(* IEC 61131-3 sources: kns-port-domestic/targets/astra/lib/src/POUs/Util/FB_StartsWindow, 7 files *)

(* ---- FB_StartsWindow.decl.st ---- *)
// Назначение: пуски за скользящий час (лимит пусков двигателя). Кольцо отметок LTIME,
//             упорядоченных по времени: самая старая — в начале, самая новая — в конце.
//             Отметки старше окна и «из будущего» (время назад) удаляются. Окно не
//             энергонезависимо: после перезапуска ПЛК оно пустое (A-03).
// Автор:      kr0nsch
// Версия:     0.1.0
// Документ:   docs/fb/FB_StartsWindow.md
FUNCTION_BLOCK FB_StartsWindow
VAR
    altStart : ARRAY[0..GVL_Const.STARTS_WINDOW_MAX - 1] OF LTIME;   // кольцо отметок пусков
    uiNext   : UINT;      // индекс следующей записи
    uiUsed   : UINT;      // занято записей, 0..STARTS_WINDOW_MAX
END_VAR

(* ---- Count.method.decl.st ---- *)
// Число отметок t с t <= ltNow и ltNow - t < STARTS_WINDOW. Отметки «из будущего» (время
// назад) и старше окна удаляются
METHOD PUBLIC Count : UINT
VAR_INPUT
    ltNow : LTIME;    // текущее время
END_VAR
VAR
    xMore : BOOL;     // продолжать удаление
    uiLast : UINT;    // индекс самой новой отметки
    uiFirst : UINT;   // индекс самой старой отметки
END_VAR

(* ---- Count.method.impl.st ---- *)
// 1. Отметки «из будущего» — с конца
xMore := uiUsed > 0;
WHILE xMore DO
    uiLast := (uiNext + GVL_Const.STARTS_WINDOW_MAX - 1) MOD GVL_Const.STARTS_WINDOW_MAX;
    IF altStart[uiLast] > ltNow THEN
        uiNext := uiLast;
        uiUsed := uiUsed - 1;
        xMore := uiUsed > 0;
    ELSE
        xMore := FALSE;
    END_IF
END_WHILE

// 2. Отметки старше окна — с начала. Все оставшиеся <= ltNow: разность без переполнения
xMore := uiUsed > 0;
WHILE xMore DO
    uiFirst := (uiNext + GVL_Const.STARTS_WINDOW_MAX - uiUsed) MOD GVL_Const.STARTS_WINDOW_MAX;
    IF ltNow - altStart[uiFirst] >= GVL_Const.STARTS_WINDOW THEN
        uiUsed := uiUsed - 1;
        xMore := uiUsed > 0;
    ELSE
        xMore := FALSE;
    END_IF
END_WHILE

Count := uiUsed;

(* ---- Register.method.decl.st ---- *)
// Добавить отметку пуска; при заполнении кольца затирается самая старая
METHOD PUBLIC Register
VAR_INPUT
    ltNow : LTIME;   // время пуска
END_VAR
VAR
    xMore : BOOL;    // продолжать удаление с конца
    uiLast : UINT;   // индекс самой новой отметки
END_VAR

(* ---- Register.method.impl.st ---- *)
// 1. Отметки новее регистрируемой (было «время назад») удаляются: кольцо остаётся упорядоченным
xMore := uiUsed > 0;
WHILE xMore DO
    uiLast := (uiNext + GVL_Const.STARTS_WINDOW_MAX - 1) MOD GVL_Const.STARTS_WINDOW_MAX;
    IF altStart[uiLast] > ltNow THEN
        uiNext := uiLast;
        uiUsed := uiUsed - 1;
        xMore := uiUsed > 0;
    ELSE
        xMore := FALSE;
    END_IF
END_WHILE

// 2. Запись; заполненное кольцо затирает самую старую отметку
altStart[uiNext] := ltNow;
uiNext := (uiNext + 1) MOD GVL_Const.STARTS_WINDOW_MAX;
uiUsed := MIN(uiUsed + 1, GVL_Const.STARTS_WINDOW_MAX);

(* ---- TimeToFree.method.decl.st ---- *)
// Через сколько число пусков в окне станет меньше uiMax; LTIME#0S, если uiMax = 0 (без
// ограничения) или пусков уже меньше uiMax
METHOD PUBLIC TimeToFree : LTIME
VAR_INPUT
    ltNow : LTIME;    // текущее время
    uiMax : UINT;     // лимит пусков в окне
END_VAR
VAR
    uiCount : UINT;   // пусков в окне
    uiIdx : UINT;     // индекс отметки, после истечения которой пусков станет uiMax - 1
END_VAR

(* ---- TimeToFree.method.impl.st ---- *)
uiCount := Count(ltNow := ltNow);
IF uiMax = 0 OR uiCount < uiMax THEN
    // PORT: [types] проверить в Astra.IDE — литералы и преобразования LTIME (C11)
    TimeToFree := LTIME#0S;
ELSE
    // отметки упорядочены: должна истечь (uiCount - uiMax)-я от самой старой (с нуля).
    // Она в окне, поэтому ltNow - t < STARTS_WINDOW и результат больше нуля
    uiIdx := (uiNext + GVL_Const.STARTS_WINDOW_MAX - uiUsed + uiCount - uiMax) MOD GVL_Const.STARTS_WINDOW_MAX;
    TimeToFree := GVL_Const.STARTS_WINDOW - (ltNow - altStart[uiIdx]);
END_IF
